(* PLC project Vn_fb_tp, Beckhoff Automation GmbH TwinCAT PLC Control 3.5.13.21 *)
(* stored: creationDateTime 1970-01-01T00:00:00 *)

PROGRAM Vn_fb_tp

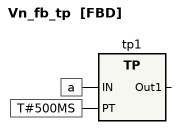
(* FBD diagram, written out as Structured Text *)
tp1(IN := a, PT := T#500MS);
END_PROGRAM
